TYPE "ST_DigitalInputOutImm"
VERSION : 0.1
   STRUCT
      "Value" : Bool;
      "Quality" : Bool;
   END_STRUCT;
END_TYPE
